(* IEC 61131-3 sources: RepoSTGen/dataset/project_code/counter/PRG, 1 file *)

(* ---- PLC_PRG.st ---- *)
PROGRAM PLC_PRG
VAR
	FB_Counter_0:FB_Counter;
	bUp,bDown,bReset:BOOL;
	ActuallyValue:int;
END_VAR

FB_Counter_0(
    bUp := bUp,
    bDown := bDown,
    bReset := bReset
);

ActuallyValue := FB_Counter_0.nValue;
